PROGRAM main
  VAR
    SCADA_HVAC_ENABLE AT %QX0.0 : BOOL;
    PUB_COMPRESSOR_RUNNING AT %QX0.1 : BOOL;
    PUB_HVAC_FAULT AT %QX0.2 : BOOL;
    SCADA_TARGET_TEMP_C AT %QW0 : UINT;
    PUB_TEMP_C AT %QW1 : UINT;
    PUB_HUMIDITY_PCT AT %QW2 : UINT;
    PUB_HEARTBEAT AT %QW3 : UINT;
    PUB_RECONNECT_COUNT AT %QW4 : UINT;
    HVAC_ENABLE AT %QX100.0 : BOOL;
    TARGET_TEMP_C AT %QW100 : UINT;
    COMPRESSOR_RUNNING AT %IX100.0 : BOOL;
    HVAC_FAULT AT %IX100.1 : BOOL;
    TEMP_C AT %IW100 : UINT;
    HUMIDITY_PCT AT %IW101 : UINT;
    HEARTBEAT AT %IW102 : UINT;
    RECONNECT_COUNT AT %IW103 : UINT;
  END_VAR

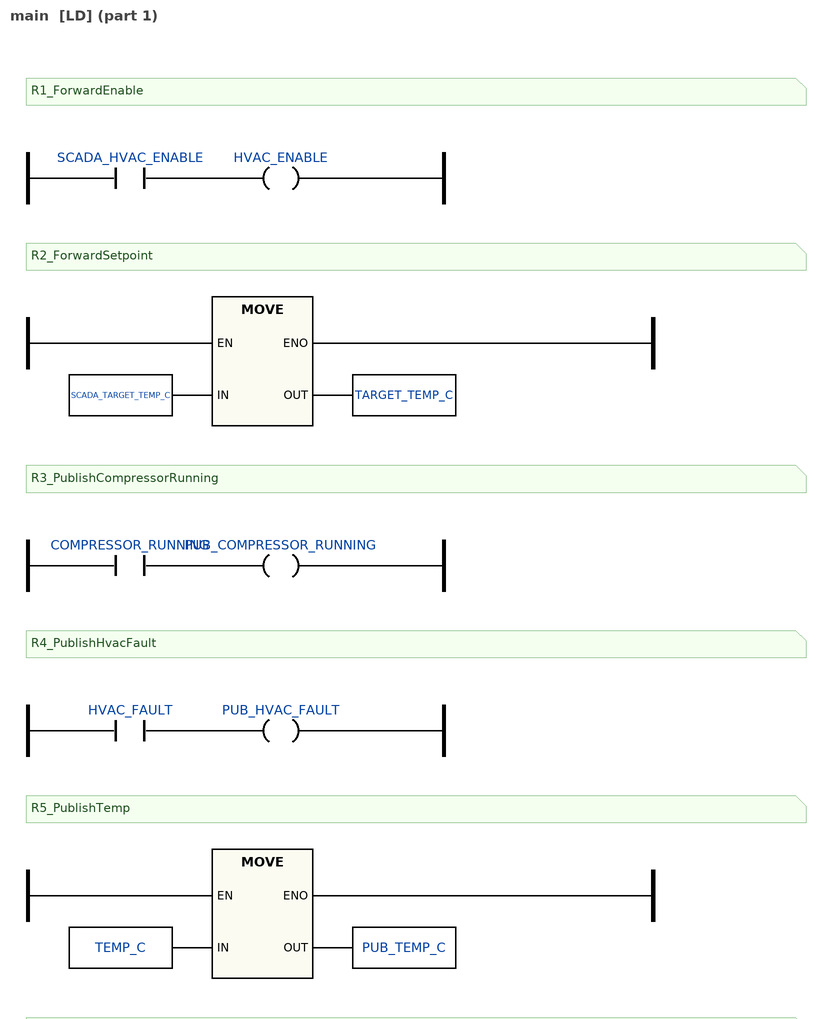
(* LD diagram, written out as Structured Text *)
(* R1_ForwardEnable *)
HVAC_ENABLE := SCADA_HVAC_ENABLE;
(* R2_ForwardSetpoint *)
TARGET_TEMP_C := SCADA_TARGET_TEMP_C;
(* R3_PublishCompressorRunning *)
PUB_COMPRESSOR_RUNNING := COMPRESSOR_RUNNING;
(* R4_PublishHvacFault *)
PUB_HVAC_FAULT := HVAC_FAULT;
(* R5_PublishTemp *)
PUB_TEMP_C := TEMP_C;
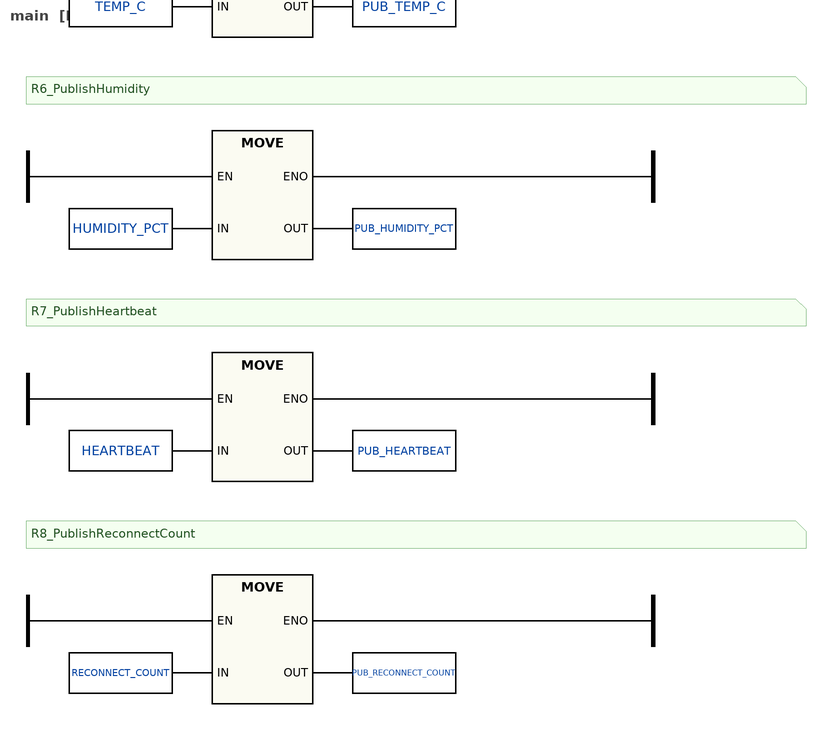
(* R6_PublishHumidity *)
PUB_HUMIDITY_PCT := HUMIDITY_PCT;
(* R7_PublishHeartbeat *)
PUB_HEARTBEAT := HEARTBEAT;
(* R8_PublishReconnectCount *)
PUB_RECONNECT_COUNT := RECONNECT_COUNT;
END_PROGRAM
